//{attribute 'qualified_only'}
VAR_GLOBAL
	stVisuPLC_To_PLC		AT %MB1000 : ST_VisuPLC_To_PLC;
	stPLC_To_VisuPLC		AT %MB2000 : ST_PLC_To_VisuPLC;
	
	q_stVisuPLC_To_PLC		AT %Q* : ST_VisuPLC_To_PLC;
	i_stPLC_To_VisuPLC		AT %I* : ST_PLC_To_VisuPLC;
END_VAR

(* stored: Version 1.1.0.1, ProductVersion 3.1.4024.15
   GVL g_HMI_Panel: Id {a228b303-e6d7-4b13-b3a1-b944c701c1f6} *)
